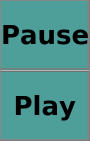
VISUALIZATION OperationButtons_1  // 90x141
VAR_IN_OUT
	stOperation	:ST_OperationButtons;
END_VAR
    Button (0,0 90x70), "Pause", colour toggle: stOperation.iActOperation=ePauseAll
        OnMouseClick: execute { stOperation.bSetPause:=TRUE; stOperation.iPauseHistory:=7; }
    Button (0,71 90x70), "Play", colour toggle: stOperation.iActOperation=ePlayAll
        OnMouseClick: execute { stOperation.bSetPlay:=TRUE; }
END_VISUALIZATION

(* stored: Version 1.1.0.1, ProductVersion 3.1.4024.13
   Visu OperationButtons_1: Id {855d9a64-56d8-4bda-b876-a7a5d053f3df} *)
